(* PLC project g_rtrig_edge, Anonymous Benchmark Suite 1.0 *)
(* stored: creationDateTime 2026-07-09T00:00:00 *)

PROGRAM g_rtrig_edge
  VAR_INPUT
    Sig : BOOL;
  END_VAR
  VAR_OUTPUT
    Rise : BOOL;
    OneShot : BOOL;
    Sig_prev : BOOL;
  END_VAR

(* LD diagram, written out as Structured Text *)
Rise := Sig AND NOT Sig_prev;
OneShot := Rise;
Sig_prev := Sig;
END_PROGRAM

CONFIGURATION Config0
  RESOURCE Res0 ON PLC
    TASK tcyclic(INTERVAL := T#10ms, PRIORITY := 0);
    PROGRAM inst0 WITH tcyclic : g_rtrig_edge;
  END_RESOURCE
END_CONFIGURATION
